FUNCTION_BLOCK FB_Safety
VAR_INPUT
END_VAR
VAR_OUTPUT
END_VAR
VAR
END_VAR

END_FUNCTION_BLOCK

(* stored: Version 1.1.0.1
   POU FB_Safety: Id {599f50d2-150a-434f-a0e9-82868f458a41}, SpecialFunc None *)
